Fanuc KAREL source: KA00151.KL

PROGRAM KA00151
%NOLOCKGROUP
VAR
  SRC: ARRAY[4] OF INTEGER
  DST: ARRAY[4] OF VECTOR
BEGIN
  DST = SRC
END KA00151
